TYPE "ST_HmiResponse"
VERSION : 0.1
   STRUCT
      AckSequence : UDInt;
      Accepted : Bool;
      Diagnostic : WString[255];
      Report : "ST_ReleaseReport";
      ConfigPage : "ST_ConfigPage";
   END_STRUCT;

END_TYPE

